Fanuc KAREL source: kc00037.KL

-- PROVISIONAL review KL for V770-1; original PC SHA256 5a65d2de2a4d62ed4d6b1d516a1c87a71311e76c5cb3e66c8fb3b5f19f1f55db
-- Incomplete behavior may be omitted. Consult companion uncertainty JSON. Do not deploy.
PROGRAM KC00037
%NOLOCKGROUP
BEGIN
  -- UNRESOLVED_PC offsets 5-29; opcodes 27,22,2A,22,22,31
  -- UNRESOLVED_PC offsets 34-38; opcodes 7F
END KC00037
